(* IEC 61131-3 sources: trust-platform/libraries/oscat/src/03_data_types, 1 file *)

(* ---- oscat_data_types.st ---- *)
(* OSCAT BASIC 3.33 data types. *)

TYPE CONSTANTS_MATH :
STRUCT
    PI : REAL := 3.141592653589793;
    PI2 : REAL := 6.283185307179586;
    PI4 : REAL := 12.566370614359173;
    PI05 : REAL := 1.570796326794897;
    PI025 : REAL := 0.785398163397448;
    PI_INV : REAL := 0.318309886183791;
    E : REAL := 2.718281828459045;
    E_INV : REAL := 0.367879441171442;
    SQ2 : REAL := 1.4142135623731;
    FACTS : ARRAY[0..12] OF DINT;
END_STRUCT
END_TYPE

TYPE CONSTANTS_PHYS :
STRUCT
    C : REAL := 299792458.0;
    E : REAL := 1.60217653E-19;
    G : REAL := 9.80665;
    T0 : REAL := -273.15;
    RU : REAL := 8.314472;
    PN : REAL := 101325.0;
END_STRUCT
END_TYPE

TYPE CONSTANTS_LANGUAGE :
STRUCT
    DEFAULT : INT := 1;
    LMAX : INT := 3;
    WEEKDAYS : ARRAY[1..3, 1..7] OF STRING[10];
    WEEKDAYS2 : ARRAY[1..3, 1..7] OF STRING[2];
    MONTHS : ARRAY[1..3, 1..12] OF STRING[10];
    MONTHS3 : ARRAY[1..3, 1..12] OF STRING[3];
    DIRS : ARRAY[1..3, 0..15] OF STRING[3];
END_STRUCT
END_TYPE

TYPE CONSTANTS_LOCATION :
STRUCT
    DEFAULT : INT := 1;
    LMAX : INT := 5;
    LANGUAGE : ARRAY[1..5] OF INT;
END_STRUCT
END_TYPE

TYPE CONSTANTS_SETUP :
STRUCT
    EXTENDED_ASCII : BOOL := TRUE;
    CHARNAMES : ARRAY[1..4] OF STRING[253];
    MTH_OFS : ARRAY[1..12] OF INT;
    DECADES : ARRAY[0..8] OF REAL;
END_STRUCT
END_TYPE

TYPE CALENDAR :
STRUCT
    UTC : DT;
    LOCAL_DT : DT;
    LOCAL_DATE : DATE;
    LOCAL_TOD : TOD;
    YEAR : INT;
    MONTH : INT;
    DAY : INT;
    WEEKDAY : INT;
    OFFSET : INT;
    DST_EN : BOOL;
    DST_ON : BOOL;
    NAME : STRING[5];
    LANGUAGE : INT;
    LONGITUDE : REAL;
    LATITUDE : REAL;
    SUN_RISE : TOD;
    SUN_SET : TOD;
    SUN_MIDDAY : TOD;
    SUN_HEIGTH : REAL;
    SUN_HOR : REAL;
    SUN_VER : REAL;
    NIGHT : BOOL;
    HOLIDAY : BOOL;
    HOLY_NAME : STRING[30];
    WORK_WEEK : INT;
END_STRUCT
END_TYPE

TYPE COMPLEX :
STRUCT
    RE : REAL;
    IM : REAL;
END_STRUCT
END_TYPE

TYPE ESR_DATA :
STRUCT
    TYP : BYTE;
    ADRESS : STRING[10];
    DS : DT;
    TS : TIME;
    DATA : ARRAY[0..7] OF BYTE;
END_STRUCT
END_TYPE

TYPE FRACTION :
STRUCT
    NUMERATOR : INT;
    DENOMINATOR : INT;
END_STRUCT
END_TYPE

TYPE HOLIDAY_DATA :
STRUCT
    NAME : STRING[30];
    DAY : SINT;
    MONTH : SINT;
    USE : SINT;
END_STRUCT
END_TYPE

TYPE REAL2 :
STRUCT
    R1 : REAL;
    RX : REAL;
END_STRUCT
END_TYPE

TYPE SDT :
STRUCT
    YEAR : INT;
    MONTH : INT;
    DAY : INT;
    WEEKDAY : INT;
    HOUR : INT;
    MINUTE : INT;
    SECOND : INT;
    MS : INT;
END_STRUCT
END_TYPE

TYPE TIMER_EVENT :
STRUCT
    TYP : BYTE;
    CHANNEL : BYTE;
    DAY : BYTE;
    START : TOD;
    DURATION : TIME;
    LAND : BYTE;
    LOR : BYTE;
    LAST : DT;
END_STRUCT
END_TYPE

TYPE VECTOR_3 :
STRUCT
    X : REAL;
    Y : REAL;
    Z : REAL;
END_STRUCT
END_TYPE
